Fanuc KAREL source: kx00021.KL

-- PROVISIONAL review KL for V940-1; original PC SHA256 6f721bad0603d7622d790ae7a3c09c1126c424d39473abafbebdb7b9e614b738
-- Incomplete behavior may be omitted. Consult companion uncertainty JSON. Do not deploy.
PROGRAM KX00021
%NOLOCKGROUP
BEGIN
  -- V9_ZERO_TABLE_METADATA_HINT layout=0001; no indexed target words; source/name/runtime held
  -- UNRESOLVED_PC offsets 5-25; opcodes 2E,22,9D,33,2E,33,35
  -- UNRESOLVED_PC offsets 30-51; opcodes 22,9D,33,2E,33,34,23
  -- UNRESOLVED_PC offsets 56-60; opcodes 7F
END KX00021
